SUBAPPLICATION logiBUS_AI_Calibrated_Subscribe_VT_Lite_OPC (* Wie logiBUS_AI_Calibrated_Subscribe_VT_OPC, fuer Sensoren mit festen Referenzwerten: Remote-Subscribe CAL/RAW/MINRAW/MAXRAW -> VT-Anzeige + CO/CS-Tasten (CALL_METHOD an die Sensor-Station). Ohne lokale Re-Publishes, ohne ZERO/SPAN. *)
  (* Standard: 61499-2; Description: Copyright (c) 2026 Meisterschulen am Ostbahnhof This program and the accompanying materials are made available under the terms of the Eclipse Public License 2.0 which is available at https://www.eclipse.org/legal/epl-2.0/ SPDX-License-Identifier: EPL-2.0 *)
  (* Version 1.0, 2026-10-17, Franz Höpfinger, Meisterschulen am Ostbahnhof, Kopie von logiBUS_AI_Calibrated_Subscribe_VT_OPC (Franz: schlanke Lib-Variante bauen, damit die Lib komplett ist) - 4x AR_M2M_Subscribe_TO_Q_OPC statt AR_M2M_Subscribe_TO_Q_Publish_OPC (keine ID_*_WRITE-Spiegel), ZeroRef/SpanRef entfallen (feste Referenzwerte auf der Sensor-Station, z.B. Fuellband-Winkel). *)
  PACKAGE MyLib::sys;
  IMPORT isobus::UT::Q::const::IDs::ID_NULL;
  IMPORT isobus::UT::io::Button::ButtonActivationCode::BT_PRESSED_LATCHED;
  IMPORT logiBUS::utils::conversion::phys::NumericObjectPool_S;
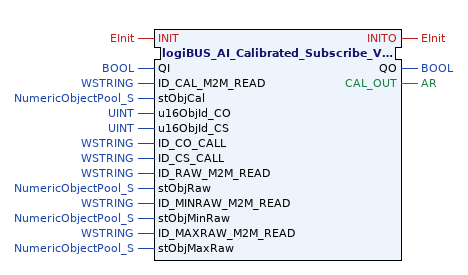
  EVENT_INPUT
    INIT : EInit; (* Initialization Request *)
  END_EVENT
  EVENT_OUTPUT
    INITO : EInit; (* Initialization Confirm *)
  END_EVENT
  VAR_INPUT
    QI : BOOL := TRUE; (* Quality Input - TRUE to enable service *)
    ID_CAL_M2M_READ : WSTRING; (* Remote-Subscribe-Adresse des kalibrierten Werts (REAL) der Sensor-Station *)
    stObjCal : logiBUS::utils::conversion::phys::NumericObjectPool_S := (u16ObjId := ID_NULL, r32Scale := 1.0, i32Offset := 0, u8Decimals := 1); (* Object ID + Scale/Offset/Decimals CNumberVariable (kalibrierter Wert) *)
    u16ObjId_CO : UINT := ID_NULL; (* Object ID Taste 'CO' (Kalibrier-Nullpunkt) auf der VT *)
    u16ObjId_CS : UINT := ID_NULL; (* Object ID Taste 'CS' (Kalibrier-Spanne) auf der VT *)
    ID_CO_CALL : WSTRING; (* Remote-Methodenadresse (CALL_METHOD) fuer den CO-Trigger auf der Sensor-Station *)
    ID_CS_CALL : WSTRING; (* Remote-Methodenadresse (CALL_METHOD) fuer den CS-Trigger auf der Sensor-Station *)
    ID_RAW_M2M_READ : WSTRING; (* Remote-Subscribe-Adresse des Rohwerts (Diagnose-Anzeige) *)
    stObjRaw : logiBUS::utils::conversion::phys::NumericObjectPool_S := (u16ObjId := ID_NULL, r32Scale := 1.0, i32Offset := 0, u8Decimals := 0); (* Object ID + Scale/Offset/Decimals CNumberVariable (Rohwert) *)
    ID_MINRAW_M2M_READ : WSTRING; (* Remote-Subscribe-Adresse Rohwert am MIN-Kalibrierpunkt (Diagnose-Anzeige) *)
    stObjMinRaw : logiBUS::utils::conversion::phys::NumericObjectPool_S := (u16ObjId := ID_NULL, r32Scale := 1.0, i32Offset := 0, u8Decimals := 0); (* Object ID + Scale/Offset/Decimals CNumberVariable (Rohwert MIN) *)
    ID_MAXRAW_M2M_READ : WSTRING; (* Remote-Subscribe-Adresse Rohwert am MAX-Kalibrierpunkt (Diagnose-Anzeige) *)
    stObjMaxRaw : logiBUS::utils::conversion::phys::NumericObjectPool_S := (u16ObjId := ID_NULL, r32Scale := 1.0, i32Offset := 0, u8Decimals := 0); (* Object ID + Scale/Offset/Decimals CNumberVariable (Rohwert MAX) *)
  END_VAR
  VAR_OUTPUT
    QO : BOOL; (* Quality Output - TRUE if service executed successfully *)
  END_VAR
  PLUGS
    CAL_OUT : adapter::types::unidirectional::AR; (* Nur-Lese-Spiegel des kalibrierten Werts fuer weitere lokale Konsumenten *)
  END_PLUGS
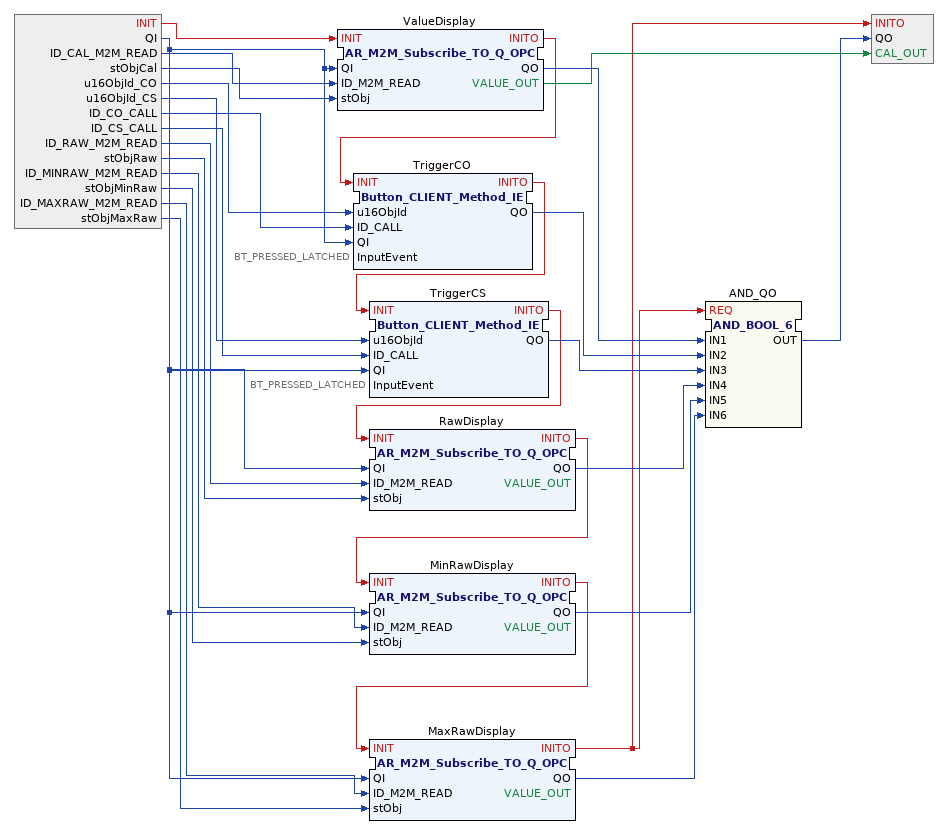
  FBS
    AND_QO : iec61131::booleanOperators::AND_BOOL_6;
  END_FBS
  SUBAPPS
    ValueDisplay : MyLib::sys::AR_M2M_Subscribe_TO_Q_OPC;
    TriggerCO : MyLib::sys::Button_CLIENT_Method_IE(InputEvent := BT_PRESSED_LATCHED);
    TriggerCS : MyLib::sys::Button_CLIENT_Method_IE(InputEvent := BT_PRESSED_LATCHED);
    RawDisplay : MyLib::sys::AR_M2M_Subscribe_TO_Q_OPC;
    MinRawDisplay : MyLib::sys::AR_M2M_Subscribe_TO_Q_OPC;
    MaxRawDisplay : MyLib::sys::AR_M2M_Subscribe_TO_Q_OPC;
  END_SUBAPPS
  EVENT_CONNECTIONS
    INIT TO ValueDisplay.INIT;
    ValueDisplay.INITO TO TriggerCO.INIT;
    TriggerCO.INITO TO TriggerCS.INIT;
    TriggerCS.INITO TO RawDisplay.INIT;
    RawDisplay.INITO TO MinRawDisplay.INIT;
    MinRawDisplay.INITO TO MaxRawDisplay.INIT;
    MaxRawDisplay.INITO TO INITO;
    MaxRawDisplay.INITO TO AND_QO.REQ;
  END_CONNECTIONS
  DATA_CONNECTIONS
    ID_CAL_M2M_READ TO ValueDisplay.ID_M2M_READ;
    stObjCal TO ValueDisplay.stObj;
    u16ObjId_CO TO TriggerCO.u16ObjId;
    u16ObjId_CS TO TriggerCS.u16ObjId;
    ID_CO_CALL TO TriggerCO.ID_CALL;
    ID_CS_CALL TO TriggerCS.ID_CALL;
    ID_RAW_M2M_READ TO RawDisplay.ID_M2M_READ;
    stObjRaw TO RawDisplay.stObj;
    ID_MINRAW_M2M_READ TO MinRawDisplay.ID_M2M_READ;
    stObjMinRaw TO MinRawDisplay.stObj;
    ID_MAXRAW_M2M_READ TO MaxRawDisplay.ID_M2M_READ;
    stObjMaxRaw TO MaxRawDisplay.stObj;
    QI TO ValueDisplay.QI;
    QI TO TriggerCO.QI;
    QI TO TriggerCS.QI;
    QI TO RawDisplay.QI;
    QI TO MinRawDisplay.QI;
    QI TO MaxRawDisplay.QI;
    ValueDisplay.QO TO AND_QO.IN1;
    TriggerCO.QO TO AND_QO.IN2;
    TriggerCS.QO TO AND_QO.IN3;
    RawDisplay.QO TO AND_QO.IN4;
    MinRawDisplay.QO TO AND_QO.IN5;
    MaxRawDisplay.QO TO AND_QO.IN6;
    AND_QO.OUT TO QO;
  END_CONNECTIONS
  ADAPTER_CONNECTIONS
    ValueDisplay.VALUE_OUT TO CAL_OUT;
  END_CONNECTIONS
END_SUBAPPLICATION
